(* IEC 61131-3 sources: daoli-st-library/DL_Process (part 64) *)

(* ---- FB_DL_ConveyorLineLink.st ---- *)
(*==============================================================================
 * 组件名称 (Component)  : FB_DL_ConveyorLineLink
 * 所属子库 (Sublibrary) : DL_Process
 * 当前版本 (Version)    : 1.0.1
 * 兼容性 (Platform)   : CODESYS 3.5 / TwinCAT 3 / 汇川 InoProShop / Machine Expert
 *                         仅依赖 Standard.library（TON / R_TRIG），零厂商方言
 * 分类     (Category)   : 工艺段功能块（Function Block · 线体级联握手协调器）
 * 功能简述 (Function)   : 相邻机台/线体段之间的级联握手协调器。把「上游有料
 *                         (BA)」「下游可收 (MR)」「强制抑制 (INH)」三类干接
 *                         点握手信号抽象为与供应商无关的状态机：三路消抖、
 *                         握手判据、传递看门狗、维护直通、同拍冲突保守侧处
 *                         理。本块只做握手编排，不直接驱动任何执行机构。
 * 首扫说明 (Init note)  : 纯事件型组件，免首扫（R23/公约 0.1），无 bInit；
 *                         所有状态由引脚沿/电平驱动，无自动首扫初始化语义。
 * 公约遵循 (Convention) : 0.2/R21 bFault 为显式排除信息级码的派生式，故障/
 *                         信息码分表标注；0.4 引脚双语同行注释；0.5/R7 全部
 *                         实例主体最前部无条件刷新，入参先算普通变量再喂实
 *                         例；0.7/R15 传递超时锁存仅复位路径清码，信息级码
 *                         瞬时型每拍重算；0.8 码位段 16#0005_xxxx（编码前经
 *                         DL_Process VERSION.md 复核：既有占用信息级
 *                         0101~0115、故障级 0200~0223，本块 0130~0133 /
 *                         0230~0231 无冲突）；0.16 无魔法数（阈值全部常量化
 *                         或引脚化）；0.17 终结符成对 ✓；0.19 码位 16# 与
 *                         【级别】同行注释；0.20 验收向量入头注释。
 * 红线自检 (Redline)    : R1 零全局变量表/外部变量引用 ✓｜R2 零物理 IO 地址 ✓
 *                         R3 纯 IEC 61131-3 ✓｜R4 看门狗/消抖/锁存复位路径 ✓
 *                         R5 全变量中英双语同行注释 ✓｜R6 ENUM+CASE+ELSE ✓
 *                         R7 六实例（R_TRIG×2/TON×4）主体最前部无条件刷新 ✓
 *                         R8 全常量化 ✓｜R25 单拍标志生命周期三律（置位-消费
 *                         -复位同周期闭环，bTransferDone 每拍先清零再置位）✓
 * 设计要点 (Key notes)  : ① 握手判据一行布尔式：上游有料(消抖 BA 或 Request)
 *                           AND 本段空 AND 下游可收 AND NOT 抑制 AND 使能
 *                           AND 无故障；同拍冲突（BA 与 Request 同真，或 MR
 *                           与 INH 同真）保守侧不放行，仅信息码暴露；
 *                         ② 传递受理 = 入口光电上升沿；料离开 = 入/出口光电
 *                           全清；完成单拍 + 计数递增；
 *                         ③ 看门狗：传递态超 tTransferTimeout → 卡料锁存
 *                           0230，仅 bReset 清；看门狗 < 消抖窗两倍自动提升
 *                           + 信息码 0133（防消抖窗吃掉整个看门狗）；
 *                         ④ 维护直通 bBypass：强制抑制输出为 FALSE 且不判超
 *                           时（信息码 0131 每拍重算）——直通会绕过卡料保护，
 *                           仅供维护调试，须审计；
 *                         ⑤ 出口断言（IF 结构保证）：向上游宣告可收与抑制上
 *                           游两输出不得同真（故障态可收输出恒 FALSE）；
 *                         ⑥ 与 FB_DL_ConveyorZone 衔接示例（仅注释，不引实
 *                           例）：本块 bMachineReadyOut → 下游区块
 *                           bDownstreamReady；下游区块 bZoneReady → 本块
 *                           bDownMachineReady。
 * 偏离留档 (Deviation)  : 依 R11 头注释留档，共 1 条：
 *                         ① eComplete「等复位」语义解释：规格未定义复位源，
 *                           按「上游 BA/Request 释放（料源已清）即视为自动复
 *                           位回 eIdle」+ bReset 手动复位双路径实现。理由：
 *                           自动线每板后手动复位不可运维；影响：eComplete 为
 *                           短暂过渡态，若调用方需强制人工确认，可不接 BA 释
 *                           放自动复位（BA 持续保持时仅 bReset 可退出）。
 * 开源溯源 (Origin)     : 来源标签 smema / conveyor-handshake（RAW_NOTES_R8
 *                         S-7：SMEMA 板级握手公开惯例——上游有料 BA、下游可
 *                         收 MR、抑制 INH 三信号电平语义与消抖/看门狗经验参
 *                         数域（消抖 20~30 ms、看门狗 5 s 量级），公开技术资
 *                         料，仅借鉴信号分类与参数域；状态机设计、码位、引脚
 *                         契约 100% 本库独立设计，clean-room 未复制任何源码。
 *                         许可证说明：SMEMA 为行业公开接口惯例，无附带许可
 *                         限制；本文件为本库原创实现，随本库许可证发布）。
 * 验收向量 (Acceptance) :
 *   V1 完整握手：BA→MR→料进（入口沿）→料出（全清）→ bTransferDone 单拍 +
 *      nTransferCount +1 → eComplete → BA 释放回 eIdle；
 *   V2 下游 INH 有效 → eInhibited，不放行，抑制解除回 eIdle + 信息码 0130；
 *   V3 传递态看门狗到 → eJamFault 锁存 0230 + bInhibitUpstream TRUE +
 *      bTransferTimeout 保持；V4 bReset 沿清锁存回 eIdle；
 *   V5 BA 与 Request 同真 → 不放行 + 信息码 0132（MR 与 INH 同真同理）；
 *   V6 bBypass 直通：bInhibitUpstream 恒 FALSE、不判超时 + 信息码 0131；
 *   V7 消抖：20 ms 毛刺（< tDebounce）被滤掉，稳定电平才参与握手；
 *   V8 故障态 bMachineReadyOut 恒 FALSE（坏料禁止放进本段）。
 * 修订历史 (Revision)   :
 *   2026-11-15  v1.0.0  首版入库（Round 08 · DL_Process 级联握手件）
 *   2026-11-15  v1.0.1  R8 总监终审修复：三路消抖 TON 的 IN 原误写为 PT 变更
 *                       掩码 _bDebBreak（常态 TRUE，三路 Q 恒 TRUE，消抖完全
 *                       失效、V7 不成立），改为「原信号 AND _bDebBreak」——原
 *                       信号为消抖对象，掩码仅承担 R14 的 PT 变更断输入一拍。
 *============================================================================*)

(*-----------------------------------------------------------------------------
 * 枚举: E_DL_LineLinkState（归属 FB_DL_ConveyorLineLink，与其同文件发布，
 *       公约 0.18 口径）。编号步长 10 留空位，eJamFault 取 99 保证排序末位
 *       （全库枚举编号惯例）。
 *----------------------------------------------------------------------------*)
TYPE E_DL_LineLinkState :
(
    eIdle         := 0,   // 空闲：无料，等上游有料信号 / Idle, no board, waiting for upstream board-available
    eBoardReady   := 10,  // 待放行：上游有料且本机可收，等下游可收 / Board ready, waiting for downstream machine-ready
    eTransferring := 20,  // 传递中：已握手，看门狗计时 / Transferring, handshake done and watchdog timing
    eComplete     := 30,  // 传递完成：料已离开本段，等复位 / Transfer complete, board left, awaiting release
    eInhibited    := 40,  // 被抑制：下游强制抑制有效，禁止启动传递 / Inhibited by downstream, transfer not allowed
    eJamFault     := 99   // 传递超时锁存：仅复位沿可退出 / Jam fault latched, only reset edge exits
) UINT;
END_TYPE

FUNCTION_BLOCK FB_DL_ConveyorLineLink
VAR_INPUT
    bEnable             : BOOL;             // 本链使能（Chain enable），FALSE=全部输出置安全侧（不放行、不请求）/ Chain enable, FALSE forces all outputs to safe side
    bUpBoardAvailable   : BOOL;             // 上游有料（Board available，上游→本机 BA 干接点），电平语义 / Upstream board available, level semantics
    bDownMachineReady   : BOOL;             // 下游可接收（Machine ready，下游→本机 MR 干接点），电平语义 / Downstream machine ready, level semantics
    bDownInhibit        : BOOL;             // 下游强制抑制（Inhibit，下游→本机 INH 干接点），TRUE=禁止放行 / Downstream inhibit, TRUE blocks release
    bBoardAtEntry       : BOOL;             // 本段入口光电（Entry photoeye），TRUE=料已进入本段 / Board present at entry photoeye
    bBoardAtExit        : BOOL;             // 本段出口光电（Exit photoeye），TRUE=料仍在本段出口 / Board present at exit photoeye
    bBoardQualityNg     : BOOL;             // 来料质量 NG 标志（Good/bad board 干接点，可选），仅透传供下游分选 / Incoming board quality NG flag, pass-through only
    bUpstreamRequest    : BOOL;             // 上游请求放料（Board requested 干接点，可选），与 BA 二选一接线 / Upstream board request, alternative to BA wiring
    tDebounce           : TIME := T#30MS;   // 输入消抖时间（Input debounce），域 T#0MS..T#1S；T#0MS=零消抖直通；经验值 20~30 ms / Input debounce time, 0 = pass-through
    tTransferTimeout    : TIME := T#5S;     // 传递看门狗（Transfer watchdog），域 T#100MS..T#60S；小于消抖窗两倍自动提升 / Transfer watchdog, auto-raised below twice debounce
    bBypass             : BOOL;             // 维护直通（Maintenance bypass），TRUE=恒放行且不报卡料，须审计，绕过卡料保护 / Maintenance bypass, overrides jam protection, audit required
    bReset              : BOOL;             // 复位超时锁存（Fault reset），上升沿受理 / Rising edge resets latched jam
END_VAR
VAR_OUTPUT
    bBoardAvailableOut  : BOOL;             // 向下游宣告有料（BA out），消抖后有料且本段已就绪 / Board available to downstream
    bMachineReadyOut    : BOOL;             // 向上游宣告可收（MR out），本段空且无故障且非抑制 / Machine ready to upstream
    bRequestBoard       : BOOL;             // 向上游请求送料（Request out），本段空且下游可收 / Board request to upstream
    bInhibitUpstream    : BOOL;             // 抑制上游（INH out），本段卡料/传递超时锁存时为 TRUE / Inhibit upstream while jammed
    bTransferring       : BOOL;             // 传递中（Transferring），传递态为 TRUE / TRUE while transferring
    bTransferDone       : BOOL;             // 传递完成单拍脉冲（Transfer done），单拍生命周期三律：每拍先清零，完成拍内置位 / One-scan transfer done pulse
    bTransferTimeout    : BOOL;             // 传递超时（Timeout），卡料锁存保持期为 TRUE / TRUE while jam latch held
    bQualityNgOut       : BOOL;             // 质量 NG 透传（NG pass-through），受理后保持下游可见直至传递完成 / NG flag held downstream-visible until complete
    bFault              : BOOL;             // 故障标志（Fault flag），显式排除信息级码（仅故障级置位）/ Fault flag, info codes excluded
    uErrorId            : UDINT;            // 故障码（Error code），16#0005_xxxx 段，0=无故障；故障级优先、无故障透出本拍信息级 / Error code, fault-level priority
    nTransferCount      : UDINT;            // 累计传递次数（Transfer counter），每完成一板 +1 / Total transfers completed
END_VAR
VAR
    _eState             : E_DL_LineLinkState := E_DL_LineLinkState.eIdle; // 内部链状态（Internal link state）/ Internal state
    _bFaultLatch        : BOOL;             // 卡料锁存标志（Jam latch flag），仅复位路径清除 / Jam latch, cleared only via reset path
    _uErrorIdInt        : UDINT;            // 内部故障级码寄存（Internal fault-level register）/ Internal fault-level register
    _uInfoCode          : UDINT;            // 本拍信息级码（Info code this cycle），瞬时型每拍重算 / Transient info code, recomputed each scan
    _bBaStable          : BOOL;             // 消抖后上游有料（Debounced BA）/ Debounced upstream board available
    _bMrStable          : BOOL;             // 消抖后下游可收（Debounced MR）/ Debounced downstream machine ready
    _bInhStable         : BOOL;             // 消抖后下游抑制（Debounced INH）/ Debounced downstream inhibit
    _bUpPresent         : BOOL;             // 归并后上游有料（Upstream present = BA 或 Request，冲突时保守侧 FALSE）/ Merged upstream present, conservative on conflict
    _bSegEmpty          : BOOL;             // 本段空（Segment empty，入口与出口光电均未遮挡）/ Segment empty by both photoeyes
    _bTransferStart     : BOOL;             // 握手判据（Transfer start condition），一行布尔式 / Transfer start handshake condition
    _bAccepted          : BOOL;             // 传递受理标志（Transfer accepted），入口光电上升沿置位 / Board accepted at entry edge
    _bNgHold            : BOOL;             // 质量 NG 保持（Quality NG hold），受理时锁存至传递完成 / Quality NG held from acceptance to completion
    _bConflict          : BOOL;             // 握手信号同拍冲突（Signal conflict this cycle），保守侧判据 / Handshake signal conflict flag
    _tWatchdogEff       : TIME := T#5S;     // 生效看门狗（Effective watchdog），被消抖窗两倍提升后的值 / Effective watchdog after auto-raise
    _tDebounceEff       : TIME := T#30MS;   // 生效消抖窗（Effective debounce），域钳位后值 / Effective debounce after clamp
    _tDebLast           : TIME := T#30MS;   // 上拍生效消抖窗（Last debounce），PT 变更检测基准 / Last debounce for PT-change detection
    _tWdLast            : TIME := T#5S;     // 上拍生效看门狗（Last watchdog），PT 变更检测基准 / Last watchdog for PT-change detection
    _bDebBreak          : BOOL := TRUE;     // 消抖输入使能（Debounce input enable），PT 变更拍断一拍 / Debounce input enable, broken on PT change
    _bWdBreak           : BOOL := TRUE;     // 看门狗输入使能（Watchdog input enable），PT 变更拍断一拍 / Watchdog input enable, broken on PT change
    _fbTonDebounceBa    : TON;              // 上游有料消抖（BA debounce timer）/ BA debounce timer
    _fbTonDebounceMr    : TON;              // 下游可收消抖（MR debounce timer）/ MR debounce timer
    _fbTonDebounceInh   : TON;              // 下游抑制消抖（INH debounce timer）/ INH debounce timer
    _fbTonWatchdog      : TON;              // 传递看门狗（Transfer watchdog timer）/ Transfer watchdog timer
    _fbTrigReset        : R_TRIG;           // 复位沿（Reset edge detector）/ Reset edge detector
    _fbTrigEntry        : R_TRIG;           // 入口光电上升沿（Entry photoeye rising edge），传递受理判据 / Entry photoedge detector
END_VAR
VAR CONSTANT
    DL_LINE_DEB_MAX     : TIME := T#1S;     // 消抖时间上限（Debounce upper clamp）/ Debounce upper clamp
    DL_LINE_WD_MIN      : TIME := T#100MS;  // 看门狗下限（Watchdog lower clamp）/ Watchdog lower clamp
    DL_LINE_WD_MAX      : TIME := T#60S;    // 看门狗上限（Watchdog upper clamp）/ Watchdog upper clamp
    DL_LINE_WD_FACTOR   : INT  := 2;        // 看门狗提升倍数（Watchdog raise factor）[-]，提升到消抖窗的此倍数 / Watchdog auto-raise factor over debounce window
    DL_LINE_ERR_JAM     : UDINT := 16#0005_0230; // 0005_0230 传递超时（卡料）【故障级】/ Transfer watchdog timeout, fault level
    DL_LINE_ERR_STATE   : UDINT := 16#0005_0231; // 0005_0231 非法状态兜底【故障级】/ Illegal state fallback, fault level
    DL_LINE_INFO_INHREL : UDINT := 16#0005_0130; // 0005_0130 下游抑制解除，恢复放行【信息级】/ Downstream inhibit released, info level
    DL_LINE_INFO_BYPASS : UDINT := 16#0005_0131; // 0005_0131 维护直通生效（每拍重算）【信息级】/ Maintenance bypass active, info level
    DL_LINE_INFO_CONFL  : UDINT := 16#0005_0132; // 0005_0132 握手信号同拍冲突（保守侧不放行）【信息级】/ Handshake signal conflict, conservative side, info level
    DL_LINE_INFO_WDRAISE: UDINT := 16#0005_0133; // 0005_0133 看门狗被提升至消抖窗两倍【信息级】/ Watchdog auto-raised to twice debounce, info level
END_VAR

// ============================================================================
// 段 1｜信息级预清零 + 实例无条件周期刷新（R7/0.5：严禁置于 IF/CASE 分支内）
//      Info preset + unconditional per-cycle refresh of all instances (R7/0.5)
// ============================================================================
_uInfoCode := 0;                        // 信息级瞬时型每拍重算（Transient info recomputed each scan）
// 消抖窗域钳位（R14：PT 变更检测先行，变更拍断输入归零 / PT change breaks input one scan）
IF tDebounce > DL_LINE_DEB_MAX THEN
    _tDebounceEff := DL_LINE_DEB_MAX;   // 超限钳位到上限（Clamped to upper bound）
ELSE
    _tDebounceEff := tDebounce;         // 引脚原值（Pin value as-is）
END_IF
// 看门狗提升值计算（R14：PT 变更检测先行 / Watchdog PT change detection first）
IF tTransferTimeout < tDebounce * DL_LINE_WD_FACTOR THEN
    _tWatchdogEff := tDebounce * DL_LINE_WD_FACTOR;      // 自动提升：防消抖窗吃掉整个看门狗（Auto-raise above debounce window）
    _uInfoCode := DL_LINE_INFO_WDRAISE; // 0005_0133 看门狗被提升【信息级】/ Watchdog raised, info level
ELSIF tTransferTimeout < DL_LINE_WD_MIN THEN
    _tWatchdogEff := DL_LINE_WD_MIN;    // 域下限钳位（Domain lower clamp）
ELSIF tTransferTimeout > DL_LINE_WD_MAX THEN
    _tWatchdogEff := DL_LINE_WD_MAX;    // 域上限钳位（Domain upper clamp）
ELSE
    _tWatchdogEff := tTransferTimeout;  // 引脚原值（Pin value as-is）
END_IF

// 三路消抖：IN 必须取「原信号」（规格 2.1-1），_bDebBreak 仅作 PT 变更拍的断输入掩码
// Three debounces: IN must be the RAW signal (spec 2.1-1); _bDebBreak is only the
// one-scan PT-change mask ANDed in, never the sole input (would make Q always TRUE)
_fbTonDebounceBa(IN := bUpBoardAvailable AND _bDebBreak, PT := _tDebounceEff);  // 上游有料消抖（BA debounce）
_fbTonDebounceMr(IN := bDownMachineReady AND _bDebBreak, PT := _tDebounceEff);  // 下游可收消抖（MR debounce）
_fbTonDebounceInh(IN := bDownInhibit AND _bDebBreak, PT := _tDebounceEff);      // 下游抑制消抖（INH debounce）
_fbTrigReset(CLK := bReset);            // 复位沿（Reset edge）
_fbTrigEntry(CLK := bBoardAtEntry);     // 入口光电沿（Entry photoedge）
_fbTonWatchdog(IN := (_eState = E_DL_LineLinkState.eTransferring) AND (NOT bBypass) AND (NOT _bWdBreak),
               PT := _tWatchdogEff);    // 传递看门狗（Transfer watchdog）

// 消抖窗/看门狗 PT 变更断输入一拍（R14：防改时间常数后计时不清零的幽灵故障）
// Debounce/watchdog PT-change one-scan input break (R14)
IF (_tDebounceEff <> _tDebLast) OR (_tWatchdogEff <> _tWdLast) THEN
    _bDebBreak := FALSE;                // 消抖输入断一拍（Debounce input broken one scan）
    _bWdBreak := FALSE;                 // 看门狗输入断一拍（Watchdog input broken one scan）
    _tDebLast := _tDebounceEff;         // 登记新消抖窗（Register new debounce）
    _tWdLast := _tWatchdogEff;          // 登记新看门狗（Register new watchdog）
ELSE
    _bDebBreak := TRUE;                 // 恢复消抖输入（Debounce input restored）
    _bWdBreak := TRUE;                  // 恢复看门狗输入（Watchdog input restored）
END_IF

// 消抖输出归并：零消抖直通（T#0MS 时 Q 有一拍滞后，此处按语义直取原信号）
// Debounce merge: pass-through raw signal when zero debounce requested
IF _tDebounceEff = T#0MS THEN
    _bBaStable := bUpBoardAvailable;    // 零消抖直通（Zero debounce pass-through）
    _bMrStable := bDownMachineReady;    // 零消抖直通（Zero debounce pass-through）
    _bInhStable := bDownInhibit;        // 零消抖直通（Zero debounce pass-through）
ELSE
    _bBaStable  := _fbTonDebounceBa.Q;  // 消抖后有料（Debounced BA）
    _bMrStable  := _fbTonDebounceMr.Q;  // 消抖后可收（Debounced MR）
    _bInhStable := _fbTonDebounceInh.Q; // 消抖后抑制（Debounced INH）
END_IF

// ============================================================================
// 段 2｜单拍标志预清零 + 复位路径（R15：锁存仅复位路径清码）
//      One-shot preset + reset path (R15)
// ============================================================================
bTransferDone := FALSE;                 // 完成单拍先清零（R25：置位-消费-复位同周期闭环）/ Done pulse preset FALSE (R25 lifecycle)

// 复位路径：仅此路径可清卡料锁存（R15）
IF _fbTrigReset.Q THEN
    _bFaultLatch := FALSE;              // 卡料锁存解除（Jam latch released）
    _uErrorIdInt := 16#0000_0000;       // 故障码清零（Fault code cleared）
END_IF

// ============================================================================
// 段 3｜派生信号与同拍冲突保守侧判定（"不猜"原则）
//      Derived signals and same-cycle conflict conservative handling
// ============================================================================
_bSegEmpty := (NOT bBoardAtEntry) AND (NOT bBoardAtExit);   // 本段空：入/出口光电均未遮挡（Segment empty）
_bConflict := (_bBaStable AND bUpstreamRequest)             // 冲突一：BA 与 Request 同真（接线错误暴露点）
           OR (_bMrStable AND _bInhStable);                 // 冲突二：MR 与 INH 同真（下游语义矛盾）
IF _bConflict THEN
    _uInfoCode := DL_LINE_INFO_CONFL;   // 0005_0132 同拍冲突，保守侧不放行【信息级】/ Conflict, conservative side, info level
END_IF
IF _bConflict OR (NOT _bBaStable) THEN
    _bUpPresent := FALSE;               // 冲突或无料 → 按无上游料处理（不猜）/ Conflict or empty means no upstream board
ELSE
    _bUpPresent := TRUE;                // 上游有料成立（Upstream board present）
END_IF

// 握手判据一行布尔式（Handshake condition, single boolean expression）：
// 上游有料 AND 本段空 AND 下游可收 AND 非抑制 AND 使能 AND 无故障 AND 无冲突
_bTransferStart := _bUpPresent AND _bSegEmpty AND _bMrStable
              AND (NOT _bInhStable) AND bEnable AND (NOT _bFaultLatch)
              AND (NOT _bConflict);

// 传递看门狗：实例已在段 1 无条件刷新（Watchdog instance refreshed unconditionally in section 1）

// ============================================================================
// 段 4｜看门狗全局监视（优先级最高，R15 锁存语义）
//      Watchdog global monitor (highest priority, latched)
// ============================================================================
IF _fbTonWatchdog.Q AND (NOT _bFaultLatch) THEN
    _bFaultLatch := TRUE;               // 传递超时锁存（Watchdog timeout latch）
    _uErrorIdInt := DL_LINE_ERR_JAM;    // 0005_0230 传递超时（卡料）【故障级】/ Transfer timeout, fault level
    _eState := E_DL_LineLinkState.eJamFault;
END_IF

// ============================================================================
// 段 5｜核心握手状态机（ENUM + CASE，含 ELSE 非法状态兜底）
//      Core handshake state machine (ENUM + CASE with ELSE fallback)
// ============================================================================
IF NOT bEnable THEN
    // 使能撤销：全部输出安全侧，状态回空闲（卡料锁存保留，仍需复位路径清）
    // Disabled: outputs to safe side, state back to idle (jam latch retained)
    _eState := E_DL_LineLinkState.eIdle;
    _bAccepted := FALSE;
ELSE
    CASE _eState OF

        E_DL_LineLinkState.eIdle: // 空闲：等上游有料
            IF _bInhStable THEN
                _eState := E_DL_LineLinkState.eInhibited;   // 下游抑制生效（Downstream inhibit active）
            ELSIF _bTransferStart THEN
                _eState := E_DL_LineLinkState.eTransferring; // 握手成立直接起传（Handshake met, start transfer）
                _bAccepted := FALSE;                         // 受理标志清零待入口沿（Accept flag armed on entry edge）
            ELSIF _bUpPresent AND _bSegEmpty AND bEnable AND (NOT _bConflict) THEN
                _eState := E_DL_LineLinkState.eBoardReady;   // 有料但下游未就绪，待放行（Board waiting for downstream ready）
            END_IF

        E_DL_LineLinkState.eBoardReady: // 待放行：等下游 MR
            IF _bInhStable THEN
                _eState := E_DL_LineLinkState.eInhibited;   // 抑制优先（Inhibit takes priority）
            ELSIF _bTransferStart THEN
                _eState := E_DL_LineLinkState.eTransferring; // 下游就绪，起传（Downstream ready, start transfer）
                _bAccepted := FALSE;
            ELSIF NOT (_bUpPresent AND _bSegEmpty) THEN
                _eState := E_DL_LineLinkState.eIdle;         // 上游料撤销或本段被占，回空闲（Upstream withdrawn or segment occupied）
            END_IF

        E_DL_LineLinkState.eTransferring: // 传递中：等受理、等料离开
            IF _fbTrigEntry.Q THEN
                _bAccepted := TRUE;              // 入口沿受理（Accepted at entry edge）
                IF bBoardQualityNg THEN
                    _bNgHold := TRUE;            // 来料 NG 锁存保持下游可见（NG held for downstream sorting）
                END_IF
            END_IF
            IF _bAccepted AND _bSegEmpty THEN
                // 料已离开本段：完成单拍 + 计数（R25：本拍内置位，段 7 出口后由下拍清零）
                // Board left: one-scan done pulse + counter increment (R25 lifecycle)
                bTransferDone := TRUE;
                nTransferCount := nTransferCount + 1;
                _eState := E_DL_LineLinkState.eComplete;
            END_IF

        E_DL_LineLinkState.eComplete: // 传递完成：等复位（偏离留档①：BA 释放自动复位 / bReset 手动复位）
            _bNgHold := FALSE;           // NG 透传随完成释放（NG pass-through released on completion）
            IF (NOT _bUpPresent) OR _fbTrigReset.Q THEN
                _eState := E_DL_LineLinkState.eIdle;     // 料源已清或手动复位（Source cleared or manual reset）
            END_IF

        E_DL_LineLinkState.eInhibited: // 被抑制：不放行
            IF NOT _bInhStable THEN
                _eState := E_DL_LineLinkState.eIdle;     // 抑制解除（Inhibit released）
                _uInfoCode := DL_LINE_INFO_INHREL;       // 0005_0130 抑制解除恢复放行【信息级】/ Inhibit released, info level
            END_IF

        E_DL_LineLinkState.eJamFault: // 卡料锁存：等复位
            IF _fbTrigReset.Q THEN
                _bAccepted := FALSE;     // 受理标志随复位清零（Accept flag cleared on reset）
            END_IF

        ELSE // 非法状态兜底（本块专用码位）
            _bFaultLatch := TRUE;        // 非法状态锁存（Illegal state latch）
            _uErrorIdInt := DL_LINE_ERR_STATE; // 0005_0231 非法状态兜底【故障级】/ Illegal state fallback, fault level
            _eState := E_DL_LineLinkState.eJamFault;
    END_CASE
END_IF

// ============================================================================
// 段 6｜输出派生（出口断言：可收输出与抑制输出不得同真）
//      Output derivation (exit assertion: ready-out and inhibit-out never both TRUE)
// ============================================================================
IF bBypass THEN
    _uInfoCode := DL_LINE_INFO_BYPASS;  // 0005_0131 维护直通生效（每拍重算）【信息级】/ Maintenance bypass active, info level
END_IF

// 向下游宣告有料：消抖后有料 + 使能 + 无故障（BA out）
bBoardAvailableOut := _bBaStable AND bEnable AND (NOT _bFaultLatch) AND (NOT _bConflict);

// 向上游宣告可收：本段空 + 使能 + 无故障 + 非抑制 + 无冲突（出口断言：故障/抑制期恒 FALSE，
// 与 bInhibitUpstream 互斥由本布尔式结构保证 / Exit assertion: mutually exclusive by construction）
bMachineReadyOut := _bSegEmpty AND bEnable AND (NOT _bFaultLatch)
               AND (NOT _bInhStable) AND (NOT _bConflict);

// 向上游请求送料：本段空 + 下游可收 + 使能 + 无故障 + 无冲突（Request out）
bRequestBoard := _bSegEmpty AND _bMrStable AND bEnable AND (NOT _bFaultLatch) AND (NOT _bConflict);

// 抑制上游：卡料锁存保持期；维护直通强制 FALSE（Inhibit upstream while jammed, voided by bypass）
bInhibitUpstream := _bFaultLatch AND (NOT bBypass);

// 状态镜像输出（State mirror outputs）
bTransferring    := (_eState = E_DL_LineLinkState.eTransferring);  // 传递中（Transferring）
bTransferTimeout := (_eState = E_DL_LineLinkState.eJamFault);      // 传递超时保持期（Timeout latch held）
bQualityNgOut    := _bNgHold;                                      // 质量 NG 透传保持（NG held visible）

// ============================================================================
// 段 7｜bFault/uErrorId 出口（R21：bFault 显式排除信息级码）
//      Outlets: bFault excludes info codes (R21)
// ============================================================================
bFault := _bFaultLatch;                 // 故障级派生式（Fault-level derived form）
IF _bFaultLatch THEN
    uErrorId := _uErrorIdInt;           // 故障级码优先透出（Fault-level priority）
ELSE
    uErrorId := _uInfoCode;             // 无故障时透出本拍信息级码（Transient info code）
END_IF
END_FUNCTION_BLOCK

(* ---- FB_DL_ConveyorZone.st ---- *)
(*==============================================================================
 * 组件名称 (Component)  : FB_DL_ConveyorZone
 * 所属子库 (Sublibrary) : DL_Process
 * 当前版本 (Version)    : 1.0.1
 * 兼容性 (Platform)   : CODESYS 3.5 / TwinCAT 3 / 汇川 InoProShop / Machine Expert
 *                         仅依赖 Standard.library（TON / R_TRIG / TP），零厂商方言
 * 分类     (Category)   : 工艺段功能块（Function Block · 输送线积放单区）
 * 功能简述 (Function)   : 单段皮带/滚筒输送线积放控制器（Zero-Pressure
 *                         Accumulation 单区）。积放单句规则：有料且下游允
 *                         许才走；卡料窗判定；run-on 清区；级联放行信号；
 *                         浪涌防护（使能沿后延迟发运行指令）；驱动控制经
 *                         I_DL_VfdDrive 接口引用（既有契约，引脚注入）。
 * 接口消费 (Consumes)   : I_DL_VfdDrive（既有接口，R6 已入库，仅引用契约文
 *                         件，零修改零新增 DUT）：运行指令 iDrive.CmdRun()/
 *                         iDrive.CmdStop()，反馈读 iDrive.bRunning/bFault。
 * 枚举归属 (Enum note)  : E_DL_ZoneState 随本块同文件发布（公约 0.11 口径：
 *                         配套枚举与主块同文件，头注释注明归属）。
 * 公约遵循 (Convention) : 0.1/R23 显式使能/指令沿驱动（无自动首扫初始化语
 *                         义），免首扫，无 bInit。
 *                         0.2/R21 bFault 显式排除信息级码；0.5/R7 全部实例
 *                         主体最前部无条件刷新；0.7/R15 卡料与故障锁存仅复
 *                         位路径清码；0.13 每拍至多一次接口方法调用。
 *                         0.8 故障码段位 16#0005_xxxx（经 DL_Process
 *                         VERSION.md 码表核对：规格建议 0005_0210/0211 已被
 *                         FB_DL_OccScheduleWindow 占用、0005_0103 已被
 *                         FB_DL_EnthalpyCompareCtrl 占用，依公约冲突顺延）：
 *                         【故障级】0005_0212 驱动指令-反馈失配、0005_0213
 *                         下游驱动故障透传、0005_0214 非法状态兜底；
 *                         【信息级】0005_0113 卡料预警（计时中未到窗）。
 * 红线自检 (Redline)    : R1 零全局变量表/外部变量引用 ✓｜R2 零物理 IO 地址 ✓
 *                         R3 纯 IEC 61131-3 ✓｜R4 时序窗防御/锁存复位路径 ✓
 *                         R5 全变量中英双语同行注释 ✓｜R6 ENUM+CASE+ELSE ✓
 *                         R7 九实例（R_TRIG×4/TON×5）主体最前部无条件刷新 ✓
 *                         R8 全常量化 ✓
 * 设计要点 (Key notes)  : ① 积放核心：RunReq = 使能 AND 无卡料 AND 无故障
 *                           AND（有料 OR 上区补跑）AND（下游允许 OR 出口空）；
 *                           末区特殊语义由调用方接线决定（bDownstreamReady
 *                           接工序就绪），本块不内判末区；
 *                         ② 驱动控制经 iDrive：RunReq 沿发 CmdRun、撤令发
 *                           CmdStop；指令-反馈失配超 tStartDelay → 故障；
 *                           方法返回 FALSE 且 iDrive.bFault → 故障透传；
 *                         ③ 卡料：RunReq 持续 + 出口光电持续遮挡超
 *                           tJamWindow → bJam 锁存（仅 bReset 清）；计时中
 *                           未到窗 → 信息级预警；
 *                         ④ 浪涌防护：使能上升沿后延迟 tStartDelay 再发运
 *                           行指令（多区级联间隔释放由各区 bZoneReady 天然
 *                           承载）；
 *                         ⑤ 手动放行：bCmdRelease 沿 → 短时放行 tRunOn
 *                           （绕过下游条件，调试用）。
 * 偏离留档 (Deviation)  : 依 R11 头注释留档，共 1 条：
 *                         ① 码位顺延：规格建议 0005_0210/0211/0103 与既有
 *                           组件冲突，依公约 0.8 顺延为 0005_0212/0213/0214
 *                           与 0005_0113（核对结果优先于建议值）。
 * 开源溯源 (Origin)     : 来源标签 conveyor-accumulation（RAW_NOTES_R7 S-9：
 *                         零积压积放（ZPA）输送线公开工程惯例——有料且下游
 *                         允许才走、run-on 清区、卡料窗、间隔释放（提取点
 *                         ⑤⑥），公开技术资料，仅借鉴规则域；状态机、接口
 *                         消费模式、码位与引脚契约 100% 本库独立设计，
 *                         clean-room 未复制源码）。
 * 验收向量 (Acceptance) :
 *   V1 有料放行/积存/清区 run-on 逐拍：bPEEntry→下游允许→运行；bPEDischarge
 *      清空后 run-on 窗停机；
 *   V2 下游阻断积放充满：bDownstreamReady=FALSE → 积存态 eAccumulating；
 *   V3 卡料窗锁存+复位：RunReq+出口遮挡超 tJamWindow → bJam + eJamFault，
 *      仅 bReset 清；
 *   V4 驱动失配：CmdRun 发出后 iDrive.bRunning 迟到超 tStartDelay → 故障
 *      0005_0212；
 *   V5 上区补跑：bUpstreamOcc=TRUE 且本区空 → 补跑合拢；
 *   V6 手动放行：bCmdRelease 沿 → tRunOn 短时放行。
 * 修订历史 (Revision)   :
 *   2026-11-15  v1.0.0  首版入库（Round 07 · DL_Process 输送线积放件）
 *   2026-11-15  v1.0.1  终审修复 2 处：① 手动放行覆盖式赋值连使能/卡料/故
 *                       障/浪涌门控一并绕过（禁用区被发出运行指令），改为仅
 *                       绕过下游条件、保留门控；② tRunOn 清区延续窗未按契
 *                       约 V1 实现（仅用于手动放行），新增 run-on 保持逻辑
 *                       （清空沿 + tRunOn 延续，使能/卡料/故障终止）
 *============================================================================*)

(*-----------------------------------------------------------------------------
 * 枚举: E_DL_ZoneState（归属 FB_DL_ConveyorZone，与其同文件）
 * 含义: 积放区状态机离散状态。编号步长 10 留空位，eJamFault 取 99 保证排
 *       序末位（全库枚举编号惯例）。
 *----------------------------------------------------------------------------*)
TYPE E_DL_ZoneState :
(
    eStopped      := 0,   // 停止：无运行指令 / Stopped, no run command
    eRunning      := 10,  // 运行：运行指令有效且驱动反馈确认 / Running, command active and drive feedback confirmed
    eAccumulating := 20,  // 积存：有料但放行条件不满足 / Accumulating, product present but release conditions unmet
    eJamFault     := 99   // 卡料/故障锁存：仅 bReset 可退出 / Jam or fault latched, only reset exits
) UINT;
END_TYPE

FUNCTION_BLOCK FB_DL_ConveyorZone
VAR_INPUT
    bPEEntry        : BOOL;             // 入口光电（Entry photoeye），TRUE=有料进入本区 / Entry photoeye, TRUE = product entering
    bPEDischarge    : BOOL;             // 出口光电（Discharge photoeye），TRUE=料仍在本区出口未清 / Discharge photoeye, TRUE = product at exit
    bDownstreamReady: BOOL;             // 下游允许放行（Downstream ready），末区接下游工序就绪；中区接下区 bZoneReady / Downstream ready, last zone ties to process ready
    bZoneEnable     : BOOL;             // 本区使能（Zone enable），FALSE=驱动停止且请求清零 / Zone enable, FALSE stops the drive
    bUpstreamOcc    : BOOL;             // 上区有料（Upstream occupied，可选过渡联动），TRUE=本区为空也补跑合拢 / Upstream occupied, gap-closing run when empty
    tRunOn          : TIME := T#1S;     // 清区延续时间（Run-on time），默认 T#1S；出口光电清空后再运行此窗 / Run-on time after the exit photoeye clears
    tJamWindow      : TIME := T#8S;     // 卡料判定窗（Jam window），默认 T#8S；按区长度/带速整定 / Jam window, tune per zone length and belt speed
    tStartDelay     : TIME := T#500MS;  // 启动确认延迟（Start feedback delay），默认 T#500MS；兼作使能沿浪涌延迟 / Start feedback delay, also the enable-edge surge delay
    bCmdRelease     : BOOL;             // 手动放行指令（Manual release，调试用），上升沿短时放行 / Manual release edge, short bypass release
    bReset          : BOOL;             // 上升沿复位卡料与故障（Reset edge clears jam and fault）/ Rising edge resets jam and fault
END_VAR
VAR_OUTPUT
    bZoneReady  : BOOL;                 // 本区就绪（Zone ready），使能无故障无卡料且本区空可接收上游来料 / Zone ready to accept upstream product
    bOccupied   : BOOL;                 // 本区有料（Zone occupied），入口或出口光电任一遮挡 / Zone occupied by either photoeye
    bJam        : BOOL;                 // 卡料锁存（Jam latched），仅 bReset 清 / Jam latched, cleared only by reset
    bFault      : BOOL;                 // 故障标志（Fault flag），显式排除信息级 / Fault flag, info codes excluded
    uErrorId    : UDINT;                // 故障码（Error code），16#0005_xxxx 段，0=无故障 / Error code, family 16#0005_xxxx
END_VAR
VAR_IN_OUT
    iDrive      : I_DL_VfdDrive;        // 本区驱动接口引用（Zone drive），由上层注入实例（既有契约 I_DL_VfdDrive）/ Zone drive interface reference injected by caller
END_VAR
VAR
    _eState        : E_DL_ZoneState := E_DL_ZoneState.eStopped; // 内部区状态（Internal zone state） / Internal state
    _bFaultLatch   : BOOL;             // 故障锁存标志（Fault latch flag），仅复位路径清除 / Fault latch, cleared only via reset path
    _uErrorIdInt   : UDINT;            // 内部故障级码寄存（Internal fault-level register）/ Internal fault-level register
    _uInfoCode     : UDINT;            // 本拍信息级码（Info code this cycle），瞬时型每拍重算 / Transient info code, recomputed each scan
    _bOccupiedInt  : BOOL;             // 内部有料派生（Internal occupied derived）/ Internal occupied derived
    _bRunReq       : BOOL;             // 积放运行请求（Accumulation run request）/ Accumulation run request
    _bRunCmdSent   : BOOL;             // 运行指令已发出锁存（Run command sent latch）/ Run command sent latch
    _bEnableDelay  : BOOL;             // 使能沿浪涌延迟激活（Enable-edge surge delay active）/ Enable-edge surge delay active
    _bManualReq    : BOOL;             // 手动放行请求（Manual release request）/ Manual release request
    _bRunOnHold    : BOOL;             // run-on 清区延续保持（Run-on sustain hold）/ Run-on sustain hold flag
    _bDriveFwd     : BOOL;             // 驱动方向登记（Drive direction registered），恒正向 / Drive direction, always forward
    _fbTrigEnable  : R_TRIG;           // 使能上升沿（Enable rising edge）/ Enable edge detector
    _fbTrigRelease : R_TRIG;           // 手动放行沿（Manual release edge）/ Manual release edge detector
    _fbTrigReset   : R_TRIG;           // 复位沿（Reset edge）/ Reset edge detector
    _fbTrigClear   : R_TRIG;           // 清空沿（Occupied falling edge），run-on 启动判据 / Occupied falling edge detector
    _fbTonJam      : TON;              // 卡料判定窗（Jam window timer）/ Jam window timer
    _fbTonFbWindow : TON;              // 指令-反馈失配窗（Command-feedback mismatch window）/ Mismatch window
    _fbTonEnable   : TON;              // 使能沿浪涌延迟（Enable-edge surge delay）/ Enable-edge surge delay
    _fbTonManual   : TON;              // 手动放行延续（Manual release sustain）/ Manual release sustain
    _fbTonRunOn    : TON;              // run-on 清区延续窗（Run-on sustain window）/ Run-on sustain window timer
END_VAR

// ============================================================================
// 段 1｜实例无条件周期刷新（R7/0.5：严禁置于 IF/CASE 分支内）
//      Unconditional per-cycle refresh of all instances (R7/0.5)
// ============================================================================
_fbTrigEnable(CLK := bZoneEnable);
_fbTrigRelease(CLK := bCmdRelease);
_fbTrigReset(CLK := bReset);
_fbTonJam(IN := _bRunReq AND bPEDischarge AND (NOT _bFaultLatch) AND (NOT bJam), PT := tJamWindow);   // 卡料窗（Jam window）
_fbTonFbWindow(IN := _bRunCmdSent XOR iDrive.bRunning, PT := tStartDelay);                            // 失配窗（Mismatch window）
_fbTonEnable(IN := _bEnableDelay, PT := tStartDelay);                                                 // 浪涌延迟（Surge delay）
_fbTonManual(IN := _bManualReq, PT := tRunOn);                                                        // 手动放行延续（Manual sustain）
_fbTrigClear(CLK := (NOT _bOccupiedInt));                                                             // 清空沿（Occupied falling edge）
_fbTonRunOn(IN := _bRunOnHold, PT := tRunOn);                                                         // run-on 清区延续窗（Run-on sustain window）

// ============================================================================
// 段 2｜信息级预清零 + 复位路径（R15：卡料与故障锁存仅复位路径清码）
//      Info preset + reset path (R15)
// ============================================================================
_uInfoCode := 0;                  // 信息级瞬时型每拍重算（Transient info recomputed each scan）

IF _fbTrigReset.Q THEN
    bJam := FALSE;                // 卡料锁存解除（Jam released）
    _bFaultLatch := FALSE;        // 故障锁存解除（Fault latch released）
    _uErrorIdInt := 16#0000_0000; // 故障码清零（Fault code cleared）
END_IF

// ============================================================================
// 段 3｜故障全局监视（优先级最高）：失配 / 驱动故障透传
//      Global fault monitors: command-feedback mismatch / drive fault pass-through
// ============================================================================
IF _fbTonFbWindow.Q AND (NOT _bFaultLatch) THEN
    _bFaultLatch := TRUE;         // 指令-反馈失配锁存（Mismatch latch）
    _uErrorIdInt := 16#0005_0212; // 0005_0212 驱动指令-反馈失配【故障级】/ Drive command-feedback mismatch, fault level
    _eState := E_DL_ZoneState.eJamFault;
END_IF
IF iDrive.bFault AND (NOT _bFaultLatch) THEN
    _bFaultLatch := TRUE;         // 下游驱动故障透传锁存（Drive fault pass-through latch）
    _uErrorIdInt := 16#0005_0213; // 0005_0213 下游驱动故障透传【故障级】/ Downstream drive fault pass-through, fault level
    _eState := E_DL_ZoneState.eJamFault;
END_IF

// ============================================================================
// 段 4｜核心积放状态机（ENUM + CASE，含 ELSE 非法状态兜底）
//      Core accumulation state machine (ENUM + CASE with ELSE fallback)
// ============================================================================
_bOccupiedInt := bPEEntry OR bPEDischarge;  // 有料派生（Occupied derived）
bOccupied := _bOccupiedInt;                 // 有料出口（Occupied outlet）

IF _fbTrigEnable.Q THEN
    _bEnableDelay := TRUE;        // 使能沿启动浪涌延迟（Enable edge arms surge delay）
END_IF
IF _fbTonEnable.Q THEN
    _bEnableDelay := FALSE;       // 浪涌延迟结束（Surge delay finished）
END_IF
IF NOT bZoneEnable THEN
    _bEnableDelay := FALSE;       // 使能撤销延迟作废（Delay voided on disable）
END_IF

IF _fbTrigRelease.Q THEN
    _bManualReq := TRUE;          // 手动放行沿登记（Manual release armed）
END_IF
IF _fbTonManual.Q THEN
    _bManualReq := FALSE;         // 手动放行延续结束（Manual sustain finished）
END_IF

// run-on 清区延续（v1.0.1 新增，契约 V1 落地）：运行中出口/入口光电全清空沿
// 启动 tRunOn 延续窗，窗内保持运行请求确保物料完全清出区段；使能撤销/卡料/
// 故障立即终止（Run-on hold: keep running tRunOn after the product clears,
// cancelled by disable/jam/fault, v1.0.1）
IF _fbTrigClear.Q AND _bRunCmdSent AND bZoneEnable AND (NOT bJam) AND (NOT _bFaultLatch) THEN
    _bRunOnHold := TRUE;          // 运行中清空沿启动延续窗（Clear edge while running arms the hold）
END_IF
IF _fbTonRunOn.Q OR (NOT bZoneEnable) OR bJam OR _bFaultLatch THEN
    _bRunOnHold := FALSE;         // 延续窗到期或门控撤销终止（Hold released on expiry or gating loss）
END_IF

// 积放单句规则：有料（或上区补跑）且下游允许（或出口空）才走（末区语义由接
// 线承担，本块不内判末区）；run-on 清区延续：出口光电清空后继续运行 tRunOn
// 窗确保完全清出（v1.0.1 按契约 V1 落地）
// ZPA rule: run when occupied (or gap-closing) AND downstream ready (or exit clear);
// run-on hold keeps the belt running tRunOn after the product clears (v1.0.1)
_bRunReq := bZoneEnable AND (NOT bJam) AND (NOT _bFaultLatch)
        AND (_bOccupiedInt OR bUpstreamOcc OR _bRunOnHold)
        AND (bDownstreamReady OR (NOT bPEDischarge))
        AND (NOT _bEnableDelay);  // 浪涌延迟未过不发令（No command before surge delay elapses）
IF _bManualReq THEN
    // 手动放行仅绕过下游条件（v1.0.1 修复：原覆盖式赋值连使能/卡料/故障/浪涌
    // 门控一并绕过，禁用区会被发出运行指令）/ Manual release bypasses the
    // downstream condition ONLY, gating preserved (v1.0.1 fix)
    _bRunReq := bZoneEnable AND (NOT bJam) AND (NOT _bFaultLatch) AND (NOT _bEnableDelay);
END_IF

IF bJam OR _bFaultLatch THEN
    CASE _eState OF
        E_DL_ZoneState.eJamFault: ; // 锁存态等待复位（Latched, awaiting reset）
        ELSE
            _eState := E_DL_ZoneState.eJamFault; // 锁存标志同步（Latch state sync）
    END_CASE
ELSIF NOT bZoneEnable THEN
    _eState := E_DL_ZoneState.eStopped; // 未使能停止（Disabled stop）
    _bRunCmdSent := FALSE;              // 撤销指令锁存（Command latch revoked）
ELSE
    CASE _eState OF

        E_DL_ZoneState.eStopped: // 停止态：评估运行请求
            IF _bRunReq THEN
                _eState := E_DL_ZoneState.eRunning; // 受理运行（Run accepted）
            END_IF

        E_DL_ZoneState.eRunning: // 运行态：撤令回停止/积存
            IF NOT _bRunReq THEN
                IF _bOccupiedInt THEN
                    _eState := E_DL_ZoneState.eAccumulating; // 有料积存（Accumulate）
                ELSE
                    _eState := E_DL_ZoneState.eStopped;      // 空区停止（Stopped when empty）
                END_IF
            END_IF

        E_DL_ZoneState.eAccumulating: // 积存态：等待放行条件
            IF _bRunReq THEN
                _eState := E_DL_ZoneState.eRunning; // 放行（Release）
            ELSIF NOT _bOccupiedInt THEN
                _eState := E_DL_ZoneState.eStopped; // 清空停止（Stopped when cleared）
            END_IF

        E_DL_ZoneState.eJamFault: // 卡料/故障态：复位路径见段 2
            IF NOT bJam THEN
                _eState := E_DL_ZoneState.eStopped; // 复位后回停止（Back to stopped after reset）
            END_IF

        ELSE
            // 非法状态兜底：任何越界枚举值强制锁存故障（Illegal state fallback）
            _bFaultLatch := TRUE;             // 故障锁存（Fault latch）
            _uErrorIdInt := 16#0005_0214;     // 0005_0214 非法状态兜底【故障级】/ Illegal state, fault level
            _eState := E_DL_ZoneState.eJamFault;
    END_CASE
END_IF

// ============================================================================
// 段 5｜驱动接口编排（0.13：每拍至多一次方法调用）+ 卡料锁存 + 信息级预警
//      Drive orchestration (max one method call per scan) + jam latch + info
// ============================================================================
IF _bRunReq AND (NOT _bRunCmdSent) THEN
    _bDriveFwd := TRUE;                                 // 方向登记恒正向（Direction always forward）
    IF NOT iDrive.CmdRun(bFwd := _bDriveFwd) THEN       // 发运行指令（Issue run command）
        IF iDrive.bFault THEN
            _bFaultLatch := TRUE;                       // 指令被拒且驱动故障：透传锁存（Rejected with drive fault: pass-through latch）
            _uErrorIdInt := 16#0005_0213;               // 0005_0213 下游驱动故障透传【故障级】/ Drive fault pass-through, fault level
            _eState := E_DL_ZoneState.eJamFault;
        END_IF
    ELSE
        _bRunCmdSent := TRUE;                           // 指令发出锁存（Command sent latch）
    END_IF
ELSIF (NOT _bRunReq) AND _bRunCmdSent THEN
    iDrive.CmdStop();                                   // 撤令停机（Issue stop command）
    _bRunCmdSent := FALSE;                              // 撤销锁存（Latch revoked）
END_IF

IF (_fbTonJam.ET > T#0S) AND _fbTonJam.IN THEN
    _uInfoCode := 16#0005_0113;   // 0005_0113 卡料预警（计时中未到窗）【信息级】/ Jam warning (timing, below window), info level
END_IF
IF _fbTonJam.Q THEN
    bJam := TRUE;                 // 卡料窗到锁存（Jam window reached, latch）
    _eState := E_DL_ZoneState.eJamFault;
END_IF

bZoneReady := bZoneEnable AND (NOT bJam) AND (NOT _bFaultLatch) AND (NOT _bOccupiedInt); // 就绪派生（Ready derived form）

// ============================================================================
// 段 6｜bFault/uErrorId 出口（R21：bFault 显式排除信息级）
//      Outlets: bFault excludes info codes (R21)
// ============================================================================
bFault := _bFaultLatch;           // 故障级派生式（Fault-level derived form）
IF _bFaultLatch THEN
    uErrorId := _uErrorIdInt;     // 故障级码优先透出（Fault-level priority）
ELSE
    uErrorId := _uInfoCode;       // 无故障时透出本拍信息级码（Transient info code）
END_IF
END_FUNCTION_BLOCK

(* ---- FB_DL_CoolingTowerFanStageSeq.st ---- *)
(*==============================================================================
 * 组件名称 (Component)  : FB_DL_CoolingTowerFanStageSeq
 * 所属子库 (Sublibrary) : DL_Process ｜ 版本 (Version) : 1.0.0 ｜ 2026-11-24
 * 兼容性   (Platform)   : CODESYS 3.5+ / TwinCAT 3 / 汇川 InoProShop / 施耐德 Machine Expert
 *                         仅依赖 IEC 61131-3 标准库（TON / R_TRIG / LIMIT / MIN / MAX），零厂商私有库
 * 功能描述 (Function)   : 冷却塔风机分级投切与主备轮换：按 nStageCmd（0..4 台）逐台启动 / 逐台停机，
 *                         级间强制间隔 tStageGap，每台启动后 tSpinUpTol 内未见运行反馈则该台
 *                         置 aFanFault 并跳过（站级不锁存，降级继续）；累计运行时长 tRunAccum
 *                         达 nLeadRotateHours 且台数稳定时做**先进后出**主用轮换（先确认新主用
 *                         起来，再停旧主用，避免瞬时欠风量）；命令 0 台 → 逐台全停。
 *                         输出 aFanRun / aFanFault 为**内部数组的状态映射**（段 5 单点出口），
 *                         迁移与出口分离，禁止在出口数组上直接做状态记忆。
 *                         **bStart = FALSE 语义（R191 二选一，本件选「降级为安全值 + 置标志」）**：
 *                         全部 aFanRun 落 FALSE 并回 eIdle（冷却塔风机不得冻结保持）。
 * 接口     (Interface)  : 输入 bEnable / bStart / bReset（上升沿）/ nStageCmd / tStageGap /
 *                         tSpinUpTol / nLeadRotateHours / nFanCnt / bFanFb[1..4]；
 *                         输出 aFanRun[1..4] / aFanFault[1..4] / nActiveCnt / nLeadIdx /
 *                         eState（E_DL_CtfPhase）/ eCause（E_DL_CtfCause）/ bError / bValid /
 *                         tRunAccum。
 * 状态迁移表 (State Transition Table)：
 *   ① eIdle → eStartup：bEnable 且 bStart 且组态闸通过且 nStageCmd ≥ 1 且无锁存；
 *      拍 N 进入（启动）/ 本拍行为：清 aFanRun / aFanFault / 台数 / 时长、主用置 1 /
 *      拍 N+1 转出至 eStartup。
 *   ② eStartup / eStageUp → 本相内逐台启动：每 tonGap.Q 单拍启动一台（间隔 tStageGap 节拍）；
 *      拍 N 进入（间隔节拍）/ 本拍行为：置 _aFanRun[idx] 与 _nPendFan / 拍 N+1 等反馈。
 *   ③ eStartup / eStageUp → eRunning：nActiveCnt ≥ nStageCmd；拍 N 进入 / 本拍行为：
 *      发信息级 eStageStable / 拍 N+1 转出至 eRunning。
 *   ④ eRunning → eStageUp：nStageCmd 增大导致 nActiveCnt < nStageCmd（拍 N 判出 / 拍 N+1 转出）。
 *   ⑤ eRunning → eStageDown：nStageCmd 减小导致 nActiveCnt > nStageCmd。
 *   ⑥ eRunning → eRotate：tRunAccum ≥ nLeadRotateHours×3600s 且 nActiveCnt = nStageCmd ≥ 1
 *      且无挂起启动（_nPendFan = 0）；本拍行为：选下一台可用风机先启动（先进）/ 拍 N+1 转出至 eRotate。
 *   ⑦ eRotate → eRunning：新主用反馈确认 → nLeadIdx := 新台、旧主用停机（后出）、
 *      tRunAccum 清零；或 tonSpin.Q（新台启动超时）→ 该台置 aFanFault、tRunAccum 清零、
 *      信息级 eFanStartTimeout，仍回 eRunning（主用不变，降级不锁存）。
 *   ⑧ eStageDown → eRunning：nActiveCnt ≤ nStageCmd；每 tonGap.Q 单拍停一台（先停非主用，
 *      取最大下标；仅剩主用时才停主用并把主用转移到仍运行的最小下标）。
 *   ⑨ eStartup / eStageUp → eFault：命令台数不可达（_nPickIdx = 0 而 nActiveCnt < nStageCmd），
 *      锁存 eStageUnreachable（段尾迁移闸，R21）。
 *   ⑩ 任一运行相 → eFault：所有已命令风机持续无反馈达 tSpinUpTol（tonNoFb.Q），
 *      锁存 eAllFansNoFeedback。
 *   ⑪ eFault → eIdle：bReset 上升沿（R_TRIG 判 .Q）且 bEnable = FALSE（可达性自证 R152：
 *      两引脚外部恒可达，R19 穷举出口）；拍 N 进入 / 本拍行为：清锁存与成因 / 拍 N+1 转出 eIdle。
 *   ⑫ ELSE（非法枚举值）→ eFault，成因 eIllegalState（R6 兜底）。
 * 边界     (Boundary)   : ① 三个 TON（tonGap / tonSpin / tonNoFb）与 tonRun、R_TRIG 一律在 CASE 外
 *                            无条件调用（R7）；tonGap / tonSpin / tonNoFb 的 IN 均含 NOT .Q 自复位项
 *                            （R188），不依赖外部沿清零；tonGap.Q 为**单拍节拍**（自复位后仅驻留
 *                            一扫描），故每拍最多投切一台，天然限速。
 *                         ② 级间节拍自进入投切相起算（首台亦等 tStageGap），工程上留出启动冲击间隔；
 *                            若需首台立即启动，请在外部把 tStageGap 设为较小值。
 *                         ③ 数组下标安全：_nFanClamp := LIMIT(1, nFanCnt, 4)，全部 FOR 与下标访问
 *                            只用定长 1..4 与 _nFanClamp，结构性无越界（R17 定长数组）。
 *                         ④ 台数累计 run 时长用 DINT 秒累加（_diRunSec，每 1s 节拍 +1），避免 TIME
 *                            加法与乘法跨型溢出；阈值 _diRotNeed := INT_TO_DINT(h)×3600（DINT 域内）。
 *                         ⑤ 无除法、无浮点比较，故无除零与容差问题（R4）。
 *                         ⑥ 零全局耦合（无 GVL / VAR_EXTERNAL / %I / %Q，R1 / R2）。
 * 码表     (Codes)      : 本件不占用全局数字码位（R297 零码位范式）；出口为 BOOL + ENUM，
 *                         enum E_DL_CtfPhase / E_DL_CtfCause 归属本文件（全库唯一属主，R264）。
 *                         信息级（0..9）永不置 bError；故障级（10 起）赋值处一律与 _bFaultLatch
 *                         三行成对（R45），故障锁存后回放至 bReset 沿（FB33-1）。
 * 分工声明 (Scope)      : 单台风机电机保护 / 变频器故障字归 DL_Device 侧驱动件；冷却塔出水温度
 *                         PID 归 FB_DL_CoolingTowerReset / 温度回路件；本件只做**台数分级投切时序
 *                         与主备轮换**，不做温度闭环。风机反馈缺失的台级降级在此件完成，
 *                         不向上层抛故障（仅不可达 / 全无反馈才锁存）。
 * 归属     (Ownership)  : E_DL_CtfPhase / E_DL_CtfCause 归属本文件（全库唯一定义，R264）。
 * 红线自检 (Redline)    : R1 ✓ 零 GVL ｜ R2 ✓ 零 %I/%Q ｜ R3 ✓ 纯 IEC ｜ R4 ✓ 无除零/无浮点比较 +
 *                         整数域闸 ｜ R5 ✓ 逐行同行双语注释 ｜ R6 ✓ 七态 ENUM + CASE + ELSE 兜底
 *                         R7 ✓ 全部 TON/R_TRIG 在 CASE 外 ｜ R8/R9 N/A（无 METHOD）｜ R10 ✓ 无构造式
 *                         转换（INT_TO_DINT / DINT_TO_TIME）｜ R14 ✓ 无 PROPERTY ｜ R15 ✓ 无保留字
 *                         撞名（aDuty 类多字母数组名）｜ R17 ✓ 定长 ARRAY[1..4] ｜ R18 ✓ bReset 用
 *                         R_TRIG 判 .Q ｜ R19 ✓ eFault 出口 = bReset 沿 + 撤使能 ｜ R20 ✓ 启动等
 *                         反馈相带 tonSpin 超时 ｜ R21 ✓ 锁存与迁相分离（段尾迁移闸）。
 * 修订历史 (Revision)   : 2026-11-24  v1.0.0  R79-B 首版
 * 验收向量 (Acceptance) :
 *   V1 nFanCnt=3、nStageCmd=2、tStageGap=T#10S、tSpinUpTol=T#15S、bFanFb 全 TRUE：
 *      bEnable=bStart=TRUE → eStartup；第 1 个 tGap 节拍 aFanRun[1]=TRUE、nActiveCnt=1；
 *      第 2 个节拍 aFanRun[2]=TRUE、nActiveCnt=2 → eRunning、nLeadIdx=1、bValid=TRUE。
 *   V2 续 V1，nStageCmd 由 2 改 0 → eStageDown，每节拍停一台（先停非主用，最大下标优先）：
 *      先停 aFanRun[2] 再停 aFanRun[1]，nActiveCnt=0、全部 aFanRun=FALSE。
 *   V3 续 V1，nStageCmd=1 且 aFanRun[1]=TRUE 而 bFanFb[1] 始终 FALSE → tSpinUpTol 后
 *      aFanFault[1]=TRUE、aFanRun[1]=FALSE、eCause=eFanStartTimeout（信息级，bError=FALSE）、
 *      随后启动第 2 台，bError 保持 FALSE（单台降级不锁存）。
 *   V4 nFanCnt=5（越界）→ eState=eFault、eCause=eBadConfig、bError=TRUE、aFanRun 全 FALSE；
 *      bReset 上升沿且 bEnable=FALSE → 回 eIdle、bError=FALSE。
 *   V5 nLeadRotateHours=1 且台数稳定于 2 台（3# 备用）：tRunAccum 达 T#1H 后 → eRotate，
 *      先启动 aFanRun[3]（先进），确认后 nLeadIdx=3 且 aFanRun[1] 停（后出），tRunAccum 清零。
 *============================================================================*)

(*-----------------------------------------------------------------------------
 * 枚举: E_DL_CtfPhase（冷却塔风机分级投切相位；eFault 为安全相，仅 bReset 沿迁出）
 *----------------------------------------------------------------------------*)
TYPE E_DL_CtfPhase :
(
    eIdle     := 0,    // 空闲：未启动，全部风机停 / Idle: not started, all fans off
    eStartup  := 10,   // 启动相：从 0 台逐台升到命令台数 / Startup: ramp fan count up to the command
    eRunning  := 20,   // 运行相：台数已达命令值，监视与轮换判 / Running: count reached, monitor and rotation check
    eStageUp  := 30,   // 加台相：命令台数增大，逐台补启动 / Stage up: command increased, add fans one by one
    eStageDown := 40,  // 减台相：命令台数减小，逐台停机 / Stage down: command decreased, stop fans one by one
    eRotate   := 50,   // 轮换相：主用先进后出换台 / Rotate: lead change with start-before-stop
    eFault    := 90    // 故障安全相：锁存成因，风机全停 / Fault safe phase: latched cause, all fans off
);
END_TYPE

(*-----------------------------------------------------------------------------
 * 枚举: E_DL_CtfCause（成因码；信息级 = 0..9，故障级 = 10 起）
 *----------------------------------------------------------------------------*)
TYPE E_DL_CtfCause :
(
    eNone           := 0,   // 信息级：无事件 / Info: no event
    eStageStable    := 1,   // 信息级：台数与命令一致 / Info: active count matches the command
    eFanUp          := 2,   // 信息级：一台已启动并确认 / Info: one fan started and confirmed
    eFanDown        := 3,   // 信息级：一台已停机 / Info: one fan stopped
    eFanStartTimeout := 4,  // 信息级：单台启动超时，该台置 aFanFault 并跳过 / Info: one fan spin-up timeout, marked faulty and skipped
    eRotateDone     := 5,   // 信息级：主用轮换完成 / Info: lead rotation completed
    eRotateSkip     := 6,   // 信息级：无可轮换风机，本次轮换取消 / Info: no rotatable fan, rotation cancelled
    eAllFansNoFeedback := 10, // 故障级：已命令风机全部无反馈 / Fault: all commanded fans report no feedback
    eStageUnreachable  := 11, // 故障级：无可用风机可达命令台数 / Fault: fan count unreachable with the available fans
    eBadConfig      := 12,  // 故障级：台数/命令/时间参数越域 / Fault: count, command or time parameter out of domain
    eIllegalState   := 13   // 故障级：非法状态枚举值 / Fault: illegal state enum value
);
END_TYPE

FUNCTION_BLOCK FB_DL_CoolingTowerFanStageSeq
VAR_INPUT
    bEnable          : BOOL := FALSE;              // 使能：FALSE 撤全部启动命令并回 eIdle / Enable, FALSE withdraws all fan commands
    bStart           : BOOL := FALSE;              // 启动（电平）：FALSE 动作全撤 / Start level, FALSE withdraws every command
    bReset           : BOOL := FALSE;              // 复位（上升沿，需同时 bEnable=FALSE）/ Reset rising edge, requires bEnable FALSE
    nStageCmd        : INT := 0;                   // 目标风机台数，有效域 0..nFanCnt [台] / Target fan count, valid domain 0..nFanCnt
    tStageGap         : TIME := T#10S;             // 级间投切间隔，域 ≥ 100ms [s] / Inter-stage gap, domain >= 100ms
    tSpinUpTol        : TIME := T#15S;             // 单台启动确认超时，域 ≥ 100ms [s] / Spin-up confirmation timeout, domain >= 100ms
    nLeadRotateHours  : INT := 0;                  // 主备轮换小时数，0 = 不轮换，域 0..1000 [h] / Lead rotation hours, 0 disables it
    nFanCnt           : INT := 2;                  // 装机风机台数，有效域 1..4 [台] / Installed fan count, valid domain 1..4
    bFanFb            : ARRAY[1..4] OF BOOL;       // 各风机运行反馈（TRUE = 在转）[#] / Per-fan running feedback, TRUE means spinning
END_VAR
VAR_OUTPUT
    aFanRun          : ARRAY[1..4] OF BOOL;        // 各风机启动命令（内部状态映射，段 5 单点出口）[#] / Per-fan run command mapped at the tail
    aFanFault        : ARRAY[1..4] OF BOOL;        // 各风机故障标记（启动超时置位，eIdle 清除）[#] / Per-fan fault flag, set on spin-up timeout
    nActiveCnt       : INT := 0;                   // 当前在运行风机台数 [台] / Number of running fans
    nLeadIdx         : INT := 0;                   // 当前主用风机下标（1 起，0 = 无）[#] / Current lead fan index, 0 means none
    eState           : E_DL_CtfPhase;              // 状态出口（段尾单点映射）[-] / State outlet mapped at the tail
    eCause           : E_DL_CtfCause;              // 成因码出口（故障期锁存回放）[-] / Cause code outlet
    bError           : BOOL;                       // 故障锁存标志 [-] / Fault latch flag
    bValid           : BOOL;                       // 时序有效回执（投切/运行相且无锁存）[-] / Sequence validity receipt
    tRunAccum        : TIME := T#0S;               // 本轮累计运行时长（供主备轮换）[s] / Accumulated run time of this round
END_VAR
VAR
    _eState          : E_DL_CtfPhase := E_DL_CtfPhase.eIdle;  // 内部相位（CASE 唯一写入目标）[-] / Internal phase
    _bFaultLatch     : BOOL := FALSE;                          // 故障锁存位（仅 bReset 沿清除）[-] / Fault latch bit
    _eCauseLatch     : E_DL_CtfCause := E_DL_CtfCause.eNone;    // 锁存成因码（FB33-1 锁存回放）[-] / Latched cause code
    _eCauseTmp       : E_DL_CtfCause := E_DL_CtfCause.eNone;    // 本拍首因中间量（段 5 用）[-] / First cause of this scan
    _bCfgOk          : BOOL := TRUE;                           // 组态域闸通过标志 [-] / Configuration gate flag
    _bResetPulse     : BOOL := FALSE;                          // bReset 上升沿快照（R18）[-] / bReset rising-edge snapshot
    _nFanClamp       : INT := 1;                               // 装机台数钳位值 1..4 [台] / Clamped installed fan count
    _nPendFan        : INT := 0;                               // 挂起待确认的启动风机下标，0 = 无 [台] / Pending fan index awaiting confirmation
    _nOldLead        : INT := 0;                               // 轮换中旧主用下标（先进后出用）[#] / Old lead index during rotation
    _nPickIdx        : INT := 0;                               // 本拍选中的风机下标，0 = 未选中 [台] / Fan index picked in this scan
    _nIdx            : INT := 1;                               // 遍历下标（FOR 专用）[台] / Loop index for FOR statements
    _aFanRun         : ARRAY[1..4] OF BOOL;                    // 内部启动命令状态数组 [#] / Internal run-command state array
    _aFanFault       : ARRAY[1..4] OF BOOL;                    // 内部风机故障状态数组 [#] / Internal fan-fault state array
    _bAnyRun         : BOOL := FALSE;                          // 存在已命令风机标志 [-] / At least one fan commanded
    _bAnyFb          : BOOL := FALSE;                          // 存在已命令且有反馈风机标志 [-] / At least one commanded fan reports feedback
    _diRunSec        : DINT := 0;                              // 运行时长秒累加（DINT 防跨型溢出）[s] / Accumulated run seconds in DINT
    _diRotNeed       : DINT := 0;                              // 轮换阈值秒数 = 小时 × 3600，0 = 不轮换 [s] / Rotation threshold in seconds
    rtReset          : R_TRIG;                                 // bReset 边沿实例（段 2 无条件调用，R18）/ bReset edge instance called unconditionally
    tonGap           : TON;                                    // 级间节拍定时器（段 2 无条件调用）/ Inter-stage tick timer called unconditionally
    tonSpin          : TON;                                    // 单台启动确认超时（段 2 无条件调用）/ Spin-up confirmation timeout called unconditionally
    tonNoFb          : TON;                                    // 全无反馈持续判（段 2 无条件调用）/ All-fans-no-feedback persistence timer
    tonRun           : TON;                                    // 运行时长 1s 累加节拍（段 2 无条件调用）/ One-second accumulation tick timer
END_VAR
VAR CONSTANT
    DL_CTF_ZERO          : INT := 0;               // 整数零基准 [-] / Integer zero base
    DL_CTF_ONE           : INT := 1;               // 整数一起始（下标与计数）[#] / Integer one base
    DL_CTF_FAN_MAX       : INT := 4;               // 风机台数上限（数组定长）[台] / Upper bound of fans, fixed array size
    DL_CTF_ROT_MAX       : INT := 1000;            // 轮换小时数上限 [h] / Upper bound of rotation hours
    DL_CTF_GAP_MIN       : TIME := T#100MS;        // 级间间隔下限 [s] / Lower bound of the inter-stage gap
    DL_CTF_TOL_MIN       : TIME := T#100MS;        // 启动确认超时下限 [s] / Lower bound of the spin-up timeout
    DL_CTF_ONESC         : TIME := T#1S;           // 一秒累加节拍 [s] / One-second accumulation tick
    DL_CTF_SEC_PER_HOUR  : DINT := 3600;           // 每小时秒数 [s/h] / Seconds per hour
    DL_CTF_ROT_ZERO      : DINT := 0;              // DINT 零基准（轮换阈值比较）[-] / DINT zero base
END_VAR

(* —— 段 1：当拍中间量预置（不清锁存 / 数组状态 / 时长累加器，FB32-1） —— *)
_bCfgOk    := TRUE;                                    // 组态闸标志复位 / Configuration gate flag reset
_eCauseTmp := E_DL_CtfCause.eNone;                      // 当拍首因复位 / Scan cause reset
_nPickIdx  := DL_CTF_ZERO;                             // 选中下标复位 / Picked index reset
_bAnyRun   := FALSE;                                   // 已命令标志复位 / Commanded flag reset
_bAnyFb    := FALSE;                                   // 有反馈标志复位 / Feedback flag reset

(* —— 段 2：入参钳位与阈值换算（整数跨型只用标准转换，R10） —— *)
_nFanClamp := LIMIT(DL_CTF_ONE, nFanCnt, DL_CTF_FAN_MAX);                 // 台数钳位 1..4，保证下标安全 / Clamp the fan count for safe indexing
_diRotNeed := INT_TO_DINT(nLeadRotateHours) * DL_CTF_SEC_PER_HOUR;        // 轮换阈值秒数（DINT 域内不溢出）/ Rotation threshold in seconds

(* —— 段 3：组态域闸（台数 / 命令 / 时间参数，R4） —— *)
IF (nFanCnt < DL_CTF_ONE) OR (nFanCnt > DL_CTF_FAN_MAX) THEN
    _bCfgOk    := FALSE;                               // 装机台数越域 / Installed fan count out of domain
    _eCauseTmp := E_DL_CtfCause.eBadConfig;            // 故障级：组态非法 / Fault: bad configuration
ELSIF (nStageCmd < DL_CTF_ZERO) OR (nStageCmd > DL_CTF_FAN_MAX) THEN
    _bCfgOk    := FALSE;                               // 命令台数越域 / Commanded fan count out of domain
    _eCauseTmp := E_DL_CtfCause.eBadConfig;            // 故障级：组态非法 / Fault: bad configuration
ELSIF nStageCmd > nFanCnt THEN
    _bCfgOk    := FALSE;                               // 命令台数超过装机台数 / Command exceeds the installed fan count
    _eCauseTmp := E_DL_CtfCause.eBadConfig;            // 故障级：组态非法 / Fault: bad configuration
ELSIF tStageGap < DL_CTF_GAP_MIN THEN
    _bCfgOk    := FALSE;                               // 级间间隔过小 / Inter-stage gap too small
    _eCauseTmp := E_DL_CtfCause.eBadConfig;            // 故障级：组态非法 / Fault: bad configuration
ELSIF tSpinUpTol < DL_CTF_TOL_MIN THEN
    _bCfgOk    := FALSE;                               // 启动确认超时过小 / Spin-up timeout too small
    _eCauseTmp := E_DL_CtfCause.eBadConfig;            // 故障级：组态非法 / Fault: bad configuration
ELSIF (nLeadRotateHours < DL_CTF_ZERO) OR (nLeadRotateHours > DL_CTF_ROT_MAX) THEN
    _bCfgOk    := FALSE;                               // 轮换小时数越域 / Rotation hours out of domain
    _eCauseTmp := E_DL_CtfCause.eBadConfig;            // 故障级：组态非法 / Fault: bad configuration
END_IF

(* —— 段 4：边沿与定时器（CASE 外无条件调用，R7；IN 均含 NOT .Q 自复位，R188） —— *)
rtReset(CLK := bReset);                                // bReset 边沿无条件刷新（R18）/ bReset edge refreshed unconditionally
_bResetPulse := rtReset.Q;                             // 边沿快照 / Edge snapshot
tonGap(IN := ((_eState = E_DL_CtfPhase.eStartup) OR (_eState = E_DL_CtfPhase.eStageUp)
              OR (_eState = E_DL_CtfPhase.eStageDown) OR (_eState = E_DL_CtfPhase.eRotate))
             AND (NOT tonGap.Q) AND (NOT _bFaultLatch),
       PT := tStageGap);                               // 投切相内周期性单拍节拍 / Periodic single-scan tick inside the staging phases
tonSpin(IN := (_nPendFan > DL_CTF_ZERO) AND (NOT tonSpin.Q) AND (NOT _bFaultLatch),
        PT := tSpinUpTol);                             // 挂起风机启动确认超时 / Spin-up timeout of the pending fan
tonRun(IN := (_eState = E_DL_CtfPhase.eRunning) AND (nActiveCnt >= DL_CTF_ONE)
       AND (NOT tonRun.Q) AND (NOT _bFaultLatch),
       PT := DL_CTF_ONESC);                            // 运行相且至少一台在转时 1s 累加（0 台不计时）/ One-second tick only while running with at least one fan
IF tonRun.Q THEN
    _diRunSec := _diRunSec + 1;                        // 运行时长 1s 累加 / Accumulate one second of run time
END_IF
(* 全无反馈判据：已命令风机中无一返回反馈（用上一拍数组状态，一拍延迟已在头注声明） *)
FOR _nIdx := 1 TO DL_CTF_FAN_MAX DO
    IF _aFanRun[_nIdx] THEN
        _bAnyRun := TRUE;                              // 存在已命令风机 / At least one fan commanded
        IF bFanFb[_nIdx] THEN
            _bAnyFb := TRUE;                           // 该台有反馈 / This fan reports feedback
        END_IF
    END_IF
END_FOR
tonNoFb(IN := _bAnyRun AND (NOT _bAnyFb) AND (NOT tonNoFb.Q) AND (NOT _bFaultLatch),
        PT := tSpinUpTol);                             // 全无反馈持续判（超时锁存故障）/ Persistence check for the total feedback loss

(* —— 段 5：状态机主体（唯一相位写入点；故障只在分支内置锁存，迁相由段 7 统一执行） —— *)
CASE _eState OF
    E_DL_CtfPhase.eIdle :
        FOR _nIdx := 1 TO DL_CTF_FAN_MAX DO
            _aFanRun[_nIdx]   := FALSE;                // 空闲：启动命令全撤 / Idle: all run commands withdrawn
            _aFanFault[_nIdx] := FALSE;                // 空闲：台级故障标志清除 / Idle: per-fan fault flags cleared
        END_FOR
        nActiveCnt := DL_CTF_ZERO;                     // 台数清零 / Active count zeroed
        _nPendFan  := DL_CTF_ZERO;                     // 挂起启动清除 / Pending start cleared
        IF bEnable AND bStart AND _bCfgOk AND (nStageCmd > DL_CTF_ZERO) AND (NOT _bFaultLatch) THEN
            nLeadIdx        := DL_CTF_ONE;             // 主用默认第 1 台 / Lead defaults to fan one
            _diRunSec       := DL_CTF_ROT_ZERO;        // 运行时长清零 / Run seconds cleared
            _nOldLead       := DL_CTF_ZERO;            // 旧主用清零 / Old lead cleared
            eCause          := E_DL_CtfCause.eNone;    // 信息级：无事件 / Info: no event
            _eState         := E_DL_CtfPhase.eStartup; // 迁移①：进入启动相 / Move to startup
        END_IF

    E_DL_CtfPhase.eStartup :
        IF (NOT bEnable) OR (NOT bStart) THEN
            FOR _nIdx := 1 TO DL_CTF_FAN_MAX DO
                _aFanRun[_nIdx] := FALSE;              // 失能：启动命令全撤 / Disabled: withdraw all commands
            END_FOR
            nActiveCnt := DL_CTF_ZERO;                 // 台数清零 / Active count zeroed
            _nPendFan  := DL_CTF_ZERO;                 // 挂起启动清除 / Pending start cleared
            eCause     := E_DL_CtfCause.eNone;         // 信息级：无事件 / Info: no event
            _eState    := E_DL_CtfPhase.eIdle;         // 回空闲相 / Back to idle
        ELSIF nActiveCnt >= nStageCmd THEN
            eCause  := E_DL_CtfCause.eStageStable;     // 迁移③：台数已达命令值 / Count reached: stable
            _eState := E_DL_CtfPhase.eRunning;         // 进入运行相 / Move to running
        ELSIF _nPendFan > DL_CTF_ZERO THEN
            IF bFanFb[_nPendFan] THEN
                _nPendFan := DL_CTF_ZERO;              // 反馈到位：清挂起 / Feedback seen: clear the pending fan
                eCause    := E_DL_CtfCause.eFanUp;     // 信息级：一台已确认 / Info: one fan confirmed
            ELSIF tonSpin.Q THEN
                _aFanRun[_nPendFan]   := FALSE;        // 启动超时：撤该台命令 / Spin-up timeout: withdraw this command
                _aFanFault[_nPendFan] := TRUE;         // 该台置故障并跳过 / Mark this fan faulty and skip it
                nActiveCnt := nActiveCnt - DL_CTF_ONE; // 台数回退（该台未起）/ Roll the count back
                _nPendFan  := DL_CTF_ZERO;             // 清挂起 / Clear the pending fan
                eCause     := E_DL_CtfCause.eFanStartTimeout; // 信息级：单台超时降级 / Info: per-fan timeout degrade
            END_IF
        ELSIF tonGap.Q THEN
            _nPickIdx := DL_CTF_ZERO;                  // 选台前复位 / Reset the pick index
            FOR _nIdx := 1 TO _nFanClamp DO
                IF (_nPickIdx = DL_CTF_ZERO) AND (NOT _aFanRun[_nIdx]) AND (NOT _aFanFault[_nIdx]) THEN
                    _nPickIdx := _nIdx;                // 取最小可启动下标（未运行且无故障）/ Lowest startable index
                END_IF
            END_FOR
            IF _nPickIdx > DL_CTF_ZERO THEN
                _aFanRun[_nPickIdx] := TRUE;           // 迁移②：发该台启动命令 / Issue the start command
                nActiveCnt := nActiveCnt + DL_CTF_ONE; // 台数 +1 / Increment the count
                _nPendFan  := _nPickIdx;               // 挂起等反馈 / Pending confirmation
                IF nActiveCnt = DL_CTF_ONE THEN
                    nLeadIdx := _nPickIdx;             // 首台即主用 / The first fan becomes the lead
                END_IF
            ELSE
                IF NOT _bFaultLatch THEN
                    _eCauseLatch := E_DL_CtfCause.eStageUnreachable; // 故障级：台数不可达 / Fault: count unreachable
                    _bFaultLatch := TRUE;              // 置故障锁存（迁相由段 7 执行，R21）/ Latch the fault, phase moved at the tail
                END_IF
            END_IF
        END_IF

    E_DL_CtfPhase.eStageUp :
        IF (NOT bEnable) OR (NOT bStart) THEN
            FOR _nIdx := 1 TO DL_CTF_FAN_MAX DO
                _aFanRun[_nIdx] := FALSE;              // 失能：启动命令全撤 / Disabled: withdraw all commands
            END_FOR
            nActiveCnt := DL_CTF_ZERO;                 // 台数清零 / Active count zeroed
            _nPendFan  := DL_CTF_ZERO;                 // 挂起启动清除 / Pending start cleared
            eCause     := E_DL_CtfCause.eNone;         // 信息级：无事件 / Info: no event
            _eState    := E_DL_CtfPhase.eIdle;         // 回空闲相 / Back to idle
        ELSIF nActiveCnt >= nStageCmd THEN
            eCause  := E_DL_CtfCause.eStageStable;     // 台数已达命令值 / Count reached: stable
            _eState := E_DL_CtfPhase.eRunning;         // 回运行相 / Back to running
        ELSIF _nPendFan > DL_CTF_ZERO THEN
            IF bFanFb[_nPendFan] THEN
                _nPendFan := DL_CTF_ZERO;              // 反馈到位：清挂起 / Feedback seen: clear the pending fan
                eCause    := E_DL_CtfCause.eFanUp;     // 信息级：一台已确认 / Info: one fan confirmed
            ELSIF tonSpin.Q THEN
                _aFanRun[_nPendFan]   := FALSE;        // 启动超时：撤该台命令 / Spin-up timeout: withdraw this command
                _aFanFault[_nPendFan] := TRUE;         // 该台置故障并跳过 / Mark this fan faulty and skip it
                nActiveCnt := nActiveCnt - DL_CTF_ONE; // 台数回退 / Roll the count back
                _nPendFan  := DL_CTF_ZERO;             // 清挂起 / Clear the pending fan
                eCause     := E_DL_CtfCause.eFanStartTimeout; // 信息级：单台超时降级 / Info: per-fan timeout degrade
            END_IF
        ELSIF tonGap.Q THEN
            _nPickIdx := DL_CTF_ZERO;                  // 选台前复位 / Reset the pick index
            FOR _nIdx := 1 TO _nFanClamp DO
                IF (_nPickIdx = DL_CTF_ZERO) AND (NOT _aFanRun[_nIdx]) AND (NOT _aFanFault[_nIdx]) THEN
                    _nPickIdx := _nIdx;                // 取最小可启动下标 / Lowest startable index
                END_IF
            END_FOR
            IF _nPickIdx > DL_CTF_ZERO THEN
                _aFanRun[_nPickIdx] := TRUE;           // 迁移②：发该台启动命令 / Issue the start command
                nActiveCnt := nActiveCnt + DL_CTF_ONE; // 台数 +1 / Increment the count
                _nPendFan  := _nPickIdx;               // 挂起等反馈 / Pending confirmation
            ELSE
                IF NOT _bFaultLatch THEN
                    _eCauseLatch := E_DL_CtfCause.eStageUnreachable; // 故障级：台数不可达 / Fault: count unreachable
                    _bFaultLatch := TRUE;              // 置故障锁存（迁相由段 7 执行，R21）/ Latch the fault, phase moved at the tail
                END_IF
            END_IF
        END_IF

    E_DL_CtfPhase.eRunning :
        IF (NOT bEnable) OR (NOT bStart) THEN
            FOR _nIdx := 1 TO DL_CTF_FAN_MAX DO
                _aFanRun[_nIdx] := FALSE;              // 失能：启动命令全撤 / Disabled: withdraw all commands
            END_FOR
            nActiveCnt := DL_CTF_ZERO;                 // 台数清零 / Active count zeroed
            _nPendFan  := DL_CTF_ZERO;                 // 挂起启动清除 / Pending start cleared
            eCause     := E_DL_CtfCause.eNone;         // 信息级：无事件 / Info: no event
            _eState    := E_DL_CtfPhase.eIdle;         // 回空闲相 / Back to idle
        ELSIF nActiveCnt < nStageCmd THEN
            eCause  := E_DL_CtfCause.eNone;            // 信息级：无事件 / Info: no event
            _eState := E_DL_CtfPhase.eStageUp;         // 迁移④：命令增大 → 加台相 / Command increased: stage up
        ELSIF nActiveCnt > nStageCmd THEN
            eCause  := E_DL_CtfCause.eNone;            // 信息级：无事件 / Info: no event
            _eState := E_DL_CtfPhase.eStageDown;       // 迁移⑤：命令减小 → 减台相 / Command decreased: stage down
        ELSIF (_diRotNeed > DL_CTF_ROT_ZERO) AND (_diRunSec >= _diRotNeed)
              AND (nActiveCnt = nStageCmd) AND (nActiveCnt >= DL_CTF_ONE) AND (_nPendFan = DL_CTF_ZERO) THEN
            _nPickIdx := DL_CTF_ZERO;                  // 候选新主用下标复位 / Candidate index reset
            FOR _nIdx := 1 TO _nFanClamp DO
                IF (_nPickIdx = DL_CTF_ZERO) AND (NOT _aFanRun[_nIdx]) AND (NOT _aFanFault[_nIdx])
                   AND (_nIdx <> nLeadIdx) THEN
                    _nPickIdx := _nIdx;                // 取下一个可用备台（最小下标）/ Next available standby fan
                END_IF
            END_FOR
            IF _nPickIdx > DL_CTF_ZERO THEN
                _nOldLead            := nLeadIdx;      // 记录旧主用 / Record the old lead
                _aFanRun[_nPickIdx]  := TRUE;          // 迁移⑥：先进 —— 先启动新主用 / Start the new lead first
                nActiveCnt           := nActiveCnt + DL_CTF_ONE; // 过渡期多一台（瞬时加台，不欠风量）/ Temporary extra fan
                _nPendFan            := _nPickIdx;     // 挂起等确认 / Pending confirmation
                eCause               := E_DL_CtfCause.eNone; // 信息级：无事件 / Info: no event
                _eState              := E_DL_CtfPhase.eRotate; // 进入轮换相 / Move to rotation
            ELSE
                _diRunSec := DL_CTF_ROT_ZERO;          // 无备台：时长清零避免每拍重试 / No standby: clear the counter
                eCause    := E_DL_CtfCause.eRotateSkip; // 信息级：轮换取消 / Info: rotation cancelled
            END_IF
        ELSE
            eCause := E_DL_CtfCause.eStageStable;      // 信息级：台数稳定 / Info: count stable
        END_IF

    E_DL_CtfPhase.eStageDown :
        IF (NOT bEnable) OR (NOT bStart) THEN
            FOR _nIdx := 1 TO DL_CTF_FAN_MAX DO
                _aFanRun[_nIdx] := FALSE;              // 失能：启动命令全撤 / Disabled: withdraw all commands
            END_FOR
            nActiveCnt := DL_CTF_ZERO;                 // 台数清零 / Active count zeroed
            _nPendFan  := DL_CTF_ZERO;                 // 挂起启动清除 / Pending start cleared
            eCause     := E_DL_CtfCause.eNone;         // 信息级：无事件 / Info: no event
            _eState    := E_DL_CtfPhase.eIdle;         // 回空闲相 / Back to idle
        ELSIF nActiveCnt <= nStageCmd THEN
            eCause  := E_DL_CtfCause.eStageStable;     // 台数已降至命令值 / Count reduced to the command
            _eState := E_DL_CtfPhase.eRunning;         // 回运行相 / Back to running
        ELSIF tonGap.Q THEN
            _nPickIdx := DL_CTF_ZERO;                  // 停机候选复位 / Stop candidate reset
            FOR _nIdx := 1 TO _nFanClamp DO
                IF _aFanRun[_nIdx] AND (_nIdx <> nLeadIdx) THEN
                    _nPickIdx := _nIdx;                // 先停非主用（取最大下标，后投先停）/ Stop non-lead first, highest index
                END_IF
            END_FOR
            IF _nPickIdx = DL_CTF_ZERO THEN
                _nPickIdx := nLeadIdx;                 // 仅剩主用时才停主用 / Only the lead remains: stop it as well
            END_IF
            IF (_nPickIdx >= DL_CTF_ONE) AND (_nPickIdx <= DL_CTF_FAN_MAX) AND _aFanRun[_nPickIdx] THEN
                _aFanRun[_nPickIdx] := FALSE;          // 迁移⑧：停该台 / Stop this fan
                nActiveCnt := nActiveCnt - DL_CTF_ONE; // 台数 -1 / Decrement the count
                eCause     := E_DL_CtfCause.eFanDown;  // 信息级：一台已停 / Info: one fan stopped
                IF _nPickIdx = nLeadIdx THEN
                    nLeadIdx := DL_CTF_ZERO;           // 主用被停：先清主用 / Lead stopped: clear it first
                    FOR _nIdx := 1 TO _nFanClamp DO
                        IF (nLeadIdx = DL_CTF_ZERO) AND _aFanRun[_nIdx] THEN
                            nLeadIdx := _nIdx;         // 主用转移到仍运行的最小下标 / Move the lead to the lowest running fan
                        END_IF
                    END_FOR
                END_IF
            END_IF
        END_IF

    E_DL_CtfPhase.eRotate :
        IF (NOT bEnable) OR (NOT bStart) THEN
            FOR _nIdx := 1 TO DL_CTF_FAN_MAX DO
                _aFanRun[_nIdx] := FALSE;              // 失能：启动命令全撤 / Disabled: withdraw all commands
            END_FOR
            nActiveCnt := DL_CTF_ZERO;                 // 台数清零 / Active count zeroed
            _nPendFan  := DL_CTF_ZERO;                 // 挂起启动清除 / Pending start cleared
            _nOldLead  := DL_CTF_ZERO;                 // 旧主用清零 / Old lead cleared
            eCause     := E_DL_CtfCause.eNone;         // 信息级：无事件 / Info: no event
            _eState    := E_DL_CtfPhase.eIdle;         // 回空闲相 / Back to idle
        ELSIF _nPendFan > DL_CTF_ZERO THEN
            IF bFanFb[_nPendFan] THEN
                nLeadIdx             := _nPendFan;     // 迁移⑦：新主用确认，交接 / New lead confirmed: hand over
                IF (_nOldLead >= DL_CTF_ONE) AND (_nOldLead <= DL_CTF_FAN_MAX) THEN
                    _aFanRun[_nOldLead] := FALSE;      // 后出：再停旧主用 / Stop the old lead afterwards
                    nActiveCnt := nActiveCnt - DL_CTF_ONE; // 过渡多出的一台回退 / Roll back the temporary extra fan
                END_IF
                _nPendFan := DL_CTF_ZERO;              // 清挂起 / Clear the pending fan
                _nOldLead := DL_CTF_ZERO;              // 清旧主用 / Clear the old lead
                _diRunSec := DL_CTF_ROT_ZERO;          // 轮换完成，时长重新累计 / Rotation done: restart the run counter
                eCause    := E_DL_CtfCause.eRotateDone; // 信息级：轮换完成 / Info: rotation completed
                _eState   := E_DL_CtfPhase.eRunning;   // 回运行相 / Back to running
            ELSIF tonSpin.Q THEN
                _aFanRun[_nPendFan]   := FALSE;        // 新主用启动超时：撤命令 / New lead spin-up timeout: withdraw
                _aFanFault[_nPendFan] := TRUE;         // 该台置故障 / Mark this fan faulty
                nActiveCnt := nActiveCnt - DL_CTF_ONE; // 过渡台数回退 / Roll back the temporary fan
                _nPendFan  := DL_CTF_ZERO;             // 清挂起 / Clear the pending fan
                _nOldLead  := DL_CTF_ZERO;             // 清旧主用（主用不变）/ Clear the old lead, keep the lead
                _diRunSec  := DL_CTF_ROT_ZERO;         // 时长清零避免每拍重试 / Clear the counter to avoid retry storms
                eCause     := E_DL_CtfCause.eFanStartTimeout; // 信息级：降级不锁存 / Info: degrade without latching
                _eState    := E_DL_CtfPhase.eRunning;  // 回运行相 / Back to running
            END_IF
        END_IF

    E_DL_CtfPhase.eFault :
        FOR _nIdx := 1 TO DL_CTF_FAN_MAX DO
            _aFanRun[_nIdx] := FALSE;                  // 故障相：启动命令全撤（安全侧）/ Fault phase: all commands withdrawn
        END_FOR
        nActiveCnt := DL_CTF_ZERO;                     // 台数清零 / Active count zeroed
        _nPendFan  := DL_CTF_ZERO;                     // 挂起启动清除 / Pending start cleared
        IF _bResetPulse AND (NOT bEnable) THEN
            _bFaultLatch := FALSE;                     // 迁移⑪：清故障锁存 / Clear the fault latch
            _eCauseLatch := E_DL_CtfCause.eNone;       // 清锁存成因 / Clear the latched cause
            eCause       := E_DL_CtfCause.eNone;       // 出口同步归零 / Outlet follows
            _diRunSec    := DL_CTF_ROT_ZERO;           // 时长清零 / Run seconds cleared
            nLeadIdx     := DL_CTF_ONE;                // 主用回默认 / Lead back to default
            _eState      := E_DL_CtfPhase.eIdle;       // 回空闲相 / Back to idle
        END_IF

ELSE
    (* 迁移⑫：非法枚举兜底（R6） *)
    IF NOT _bFaultLatch THEN
        _eCauseLatch := E_DL_CtfCause.eIllegalState;   // 故障级：非法状态 / Fault: illegal state
        _bFaultLatch := TRUE;                          // 置故障锁存 / Latch the fault
    END_IF
END_CASE

(* —— 段 6：全无反馈持续判与组态闸的锁存（锁存与迁相分离，R21） —— *)
IF tonNoFb.Q AND (NOT _bFaultLatch) THEN
    _eCauseLatch := E_DL_CtfCause.eAllFansNoFeedback;  // 故障级：全无反馈 / Fault: total feedback loss
    _bFaultLatch := TRUE;                              // 置故障锁存 / Latch the fault
END_IF
IF (NOT _bCfgOk) AND (NOT _bFaultLatch) THEN
    _eCauseLatch := _eCauseTmp;                        // 锁存首因（组态闸）/ Latch the configuration cause
    _bFaultLatch := TRUE;                              // 置故障锁存 / Latch the fault
END_IF

(* —— 段 7：段尾故障迁移闸 + 故障相动作全撤（FB50-1④） —— *)
IF _bFaultLatch AND (_eState <> E_DL_CtfPhase.eFault) THEN
    _eState := E_DL_CtfPhase.eFault;                   // 锁存即迁相 / Latch forces the fault phase
END_IF
IF _eState = E_DL_CtfPhase.eFault THEN
    FOR _nIdx := 1 TO DL_CTF_FAN_MAX DO
        _aFanRun[_nIdx] := FALSE;                      // 故障相动作全撤（含同拍迁入）/ All commands withdrawn in fault
    END_FOR
    nActiveCnt := DL_CTF_ZERO;                         // 台数清零 / Active count zeroed
    _nPendFan  := DL_CTF_ZERO;                         // 挂起启动清除 / Pending start cleared
END_IF

(* —— 段 8：统一出口（状态映射 + 数组单点出口 + 锁存回放） —— *)
eState := _eState;                                     // 相位映射 / Phase mapping
FOR _nIdx := 1 TO DL_CTF_FAN_MAX DO
    aFanRun[_nIdx]   := _aFanRun[_nIdx];               // 启动命令映射 / Run command mapping
    aFanFault[_nIdx] := _aFanFault[_nIdx];             // 台级故障映射 / Per-fan fault mapping
END_FOR
tRunAccum := DINT_TO_TIME(_diRunSec);                  // 时长秒 → TIME（显式标准转换）/ Seconds to TIME via the standard converter
bError := _bFaultLatch;                                // 故障标志取锁存位 / Fault flag from the latch
IF _bFaultLatch THEN
    eCause := _eCauseLatch;                            // 故障期回放锁存码（FB33-1）/ Replay the latched code
END_IF
bValid := ((_eState = E_DL_CtfPhase.eRunning) OR (_eState = E_DL_CtfPhase.eStartup)
           OR (_eState = E_DL_CtfPhase.eStageUp) OR (_eState = E_DL_CtfPhase.eStageDown)
           OR (_eState = E_DL_CtfPhase.eRotate)) AND (NOT _bFaultLatch);   // 投切/运行相且无锁存时有效
END_FUNCTION_BLOCK
